(* IEC 61131-3 sources: plc-workbench/experiments/formal_r7/fault_injection/interlocked_start, 3 files *)

(* ---- before.st ---- *)
FUNCTION_BLOCK InterlockedStart
VAR_INPUT
  start : BOOL;
  stop : BOOL;
  permit : BOOL;
END_VAR
VAR_OUTPUT
  running : BOOL;
END_VAR
VAR
  prevStart : BOOL;
  startEdge : BOOL;
END_VAR
VAR WB_FaultScan : USINT; END_VAR

startEdge := start AND NOT prevStart;
prevStart := start;

IF stop OR NOT permit THEN
  running := FALSE;
ELSIF startEdge THEN
  running := TRUE;
END_IF;

WB_FaultScan := WB_FaultScan + 1;
IF WB_FaultScan = 24 THEN running := TRUE; END_IF;
END_FUNCTION_BLOCK

(* ---- candidate_01.st ---- *)
FUNCTION_BLOCK InterlockedStart
VAR_INPUT
  start : BOOL;
  stop : BOOL;
  permit : BOOL;
END_VAR
VAR_OUTPUT
  running : BOOL;
END_VAR
VAR
  prevStart : BOOL;
  startEdge : BOOL;
END_VAR

(* Edge detection uses previous scan value; block initial prevStart = FALSE *)
startEdge := start AND NOT prevStart;
prevStart := start;

(* Stop / interlock dominate any simultaneous start edge *)
IF stop OR NOT permit THEN
  running := FALSE;
ELSIF startEdge THEN
  running := TRUE;
END_IF;

END_FUNCTION_BLOCK

(* ---- candidate_final.st ---- *)
FUNCTION_BLOCK InterlockedStart
VAR_INPUT
  start : BOOL;
  stop : BOOL;
  permit : BOOL;
END_VAR
VAR_OUTPUT
  running : BOOL;
END_VAR
VAR
  prevStart : BOOL;
  startEdge : BOOL;
END_VAR

(* Edge detection uses previous scan value; block initial prevStart = FALSE *)
startEdge := start AND NOT prevStart;
prevStart := start;

(* Stop / interlock dominate any simultaneous start edge *)
IF stop OR NOT permit THEN
  running := FALSE;
ELSIF startEdge THEN
  running := TRUE;
END_IF;

END_FUNCTION_BLOCK
